// TIA Portal V21 export
// export: Created 2026-11-07T14:35:59.2461547Z, ExportSetting WithDefaults, DisplayName Totally Integrated Automation Portal, DisplayVersion V21, DisplayName STEP 7 Professional, DisplayVersion V21, DisplayName STEP 7 Safety, DisplayVersion V21, DisplayName Tech WebApplication, DisplayVersion V21, DisplayName WinCC Basic/Comfort/Advanced, DisplayVersion V21, DisplayName WinCC Unified, DisplayVersion V21
Screen "T08_Bar"  1024x768, Number=28
  ScreenLayer 
    Bar "P_Bar" at 0,0 size 100x30  CountSubDivisions=5, IntegerDigits=3, LargeTickLabelingStep=1, MaximumValue=24, Precision=2, StyleItem=Bar
      ProcessValue := BalL
